Yaskawa INFORM job: 20210126fengjipaifengkou.JBI

/JOB
//NAME 20210126fengjipaifengkou
//POS
///NPOS 7,0,0,0,0,0
///TOOL 1
///POSTYPE PULSE
///PULSE
C00000=53633,37661,-15027,0,-49471,23935
C00001=28551,52709,10228,-1332,-56280,-3343
C00002=12021,7891,-57986,977,-35407,-41870
C00003=12021,7891,-57986,977,-35407,-41870
C00004=12021,7891,-57986,977,-35407,-41870
C00005=45155,-6272,-73239,-1936,-41576,-94391
C00006=56671,33000,-22918,6788,-42680,17539
//INST
///DATE 2021/01/26 16:03
///ATTR SC,RW
///GROUP1 RB1
NOP
MOVC C00000 V=50.0
MOVC C00001 V=50.0
MOVC C00002 V=50.0
MOVC C00003 V=50.0
MOVC C00004 V=50.0
MOVC C00005 V=50.0
MOVC C00006 V=50.0
END
